{attribute 'linkalways'}
{attribute 'no_explicit_call' := 'This FB is a CLASS and must be accessed using methods or properties'}
{attribute 'enable_dynamic_creation'}
FUNCTION_BLOCK Node_F_VN_MultiplyWithContainerElements2 EXTENDS VisionNode
VAR
    ipContainer : _ITcVnContainer;
    ipDestContainer : _ITcVnContainer;
    aValue : _TcVnVector2_LREAL;
    hrPrev : _HRESULT(S_OK);
    hresult : _HRESULT(S_OK);
END_VAR

METHOD PUBLIC Clone : I_Node
VAR
    pNode : POINTER TO Node_F_VN_MultiplyWithContainerElements2;
END_VAR
pNode := __NEW(Node_F_VN_MultiplyWithContainerElements2);
Clone := pNode^;
END_METHOD

METHOD FB_init : BOOL
VAR_INPUT
    bInitRetains : BOOL;
    bInCopyCode : BOOL;
END_VAR
AddInput('ipContainer', ipContainer);
AddParameter('aValue', aValue);
AddInput('hrPrev', hrPrev);
AddOutput('ipDestContainer', ipDestContainer);
AddOutput('hresult', hresult);
END_METHOD

METHOD PROTECTED OnExecute
// The API edits the container in place. Edit a copy so the upstream container is only read.
hresult.Value := F_VN_CopyContainer(
    ipSrcContainer := ipContainer.Value,
    ipDestContainer := ipDestContainer.Value,
    hrPrev := hrPrev.Value);

hresult.Value := F_VN_MultiplyWithContainerElements2(
    aValue := aValue.Value,
    ipContainer := ipDestContainer.Value,
    hrPrev := hresult.Value);
END_METHOD

METHOD PUBLIC PreExecutionCheck
VAR_INPUT
    Check : I_PreExecutionChecks;
END_VAR
VAR
    typeGuid : GUID;
    dimensions : UINT;
END_VAR
Check.IsTrue(ipContainer.IsValid, 'ipContainer must be a valid container');
IF ipContainer.IsValid THEN
    ipContainer.Value.GetTypeGuid(typeGuid);
END_IF
dimensions := GetContainerTypeDimensions(typeGuid);
Check.IsTrue(dimensions = 2, 'ipContainer must hold TcVnPoint2 or TcVnVector2 elements');
END_METHOD

END_FUNCTION_BLOCK

(* stored: Version 1.1.0.1, ProductVersion 3.1.4026.19
   POU Node_F_VN_MultiplyWithContainerElements2: Id {2f8cc159-7fda-4abf-955b-89e0e17bf5c9}, SpecialFunc None
   Folder Constructor: Id {66e9e92b-8bf8-49a8-9e71-7d824c54811c}
   Method Clone: Id {a02eb8a9-975f-4187-987f-6a378660e28b}
   Method FB_init: Id {d1f6a714-8636-4409-b48e-4b83024445e0}
   Method OnExecute: Id {87c2728b-1bad-4625-b5cf-a0039c497ef3}
   Method PreExecutionCheck: Id {654bb8dd-5efe-479d-93dd-9565a256d155} *)
